Staubli VAL3: progItem.pjx

--- progItem.pjx ---
Parameters version=s8.10.3Cs9_BS2093 stackSize=5000 millimeterUnit=true
Program file=start.pgx
Program file=stop.pgx
Data file=progItem.dtx
Type name=progTemplate path=Disk://source/template/progTemplate/progTemplate.pjx

--- progItem.dtx ---
public progTemplate pProgTemplate
  [0]
    string sTRAJname
    num nType
    ifItem iIfItem
      [0]
        num nSigType[3]
        num nSigIndex[3]
        num nValue[3]
        bool bANDOR[2]
    switchItem sSwitchItem
      [0]
        num nSwitchValue
        string sIOValue
        bool bIOdisable
    forItem fForItem
      [0]
        num nLoopValue
        bool bIOdisable
        string sIOindex
        string sForTRAJ

--- start.pgx ---
program start()
begin
end

--- stop.pgx ---
program stop()
begin
end
